(* IEC 61131-3 sources: Elmo_Master/Lasal_PRG/Elmo_EtherCAT_Test_4Axis/Class/ECAT_Slave_Base (part 2) *)

        sSDOData.Buffer.pSDOCallback$^VirtualBase^.NewInst(#UserPara, #UserResult);
      end_if;

//*******************************************************************************************************************************************************
  end_case;

END_FUNCTION

FUNCTION VIRTUAL GLOBAL ECAT_Slave_Base::ClassState::NewInst
	VAR_INPUT
		pPara 	: ^CmdStruct;
		pResult 	: ^Results;
	END_VAR
	VAR_OUTPUT
		ret_code 	: IprStates;
	END_VAR
  VAR
    TmpRetCode : iprStates;
    pNewElement   : t_pHWCGetHardwareDiagnosisOutDynExt;
    pTemp : ^void;
  END_VAR

  //Return with error if command is unknown or not supported
  ret_code := ERROR;

  case pPara^.uiCmd of

//**********************************************************************************************************************************************************
    ECAT_M_SET_SLAVE_INFO:

      pResult^.uiLng := 4;
      pResult^.aData[0]$DINT := ECAT_RETERR_CMD_VERSION;

      //Check version number
      if pPara^.aPara[0]$DINT = 1 then

        pResult^.uiLng := 8;
        pResult^.aData[0]$DINT := ECAT_RETERR_CMD_PARAMETER;
        pResult^.aData[4]$DINT := 1;  //Return version number

        pSlaveInfo := pPara^.aPara[1]$^t_st_eceni_slv_info;

        //Check for valid pointer
        if pSlaveInfo then

          ret_code := READY;

          //Show slave info data on server
          DeviceAdress  := pSlaveInfo^.physaddr;
          VendorID      := pSlaveInfo^.vendorid;
          SerialNo      := pSlaveInfo^.serialno;
          ProductCode   := pSlaveInfo^.productcode;
          RevisionNo    := pSlaveInfo^.revisionno;

          pResult^.aData[0]$DINT := ECATM_OK;

          if pSlaveInfo^.name then
            DeviceNameStr.WriteDataOff(udLen:=_StrLen(pSlaveInfo^.name), udOff:=0, pData:=pSlaveInfo^.name);
          else
            LogValue("@059A (ECAT_Slave_Base::ClassState::NewInst) Invalid name in Slave-info data of Slave 0x{0}",SlaveIndex);
          end_if;

          if pSlaveInfo^.productrev then
            ProductRevStr.WriteDataOff(udLen:=_StrLen(pSlaveInfo^.productrev), udOff:=0, pData:=pSlaveInfo^.productrev);
          else
            LogValue("@059B (ECAT_Slave_Base::ClassState::NewInst) Invalid product revision in Slave-info data of Slave 0x{0}",SlaveIndex);
          end_if;
        else

        end_if;
      else
        LogError("@059C (ECAT_Slave_Base::ClassState::NewInst) Unsupported NewInst version ECAT_M_SET_SLAVE_INFO");
        ret_code := ERROR;
      end_if;

//**********************************************************************************************************************************************************
    ECAT_M_GET_SLAVE_CYCIDX:

      pResult^.uiLng := 4;
      pResult^.aData[0]$DINT := ECAT_RETERR_CMD_VERSION;

      //Check version number
      if pPara^.aPara[0]$DINT = 1 then

        pResult^.uiLng := 8;
        pResult^.aData[4]$DINT := 1;  //Return version number

        pResult^.aData[0]$DINT := ECAT_RETERR_CMD_WRONG_SLV_STATE;
        if us_InitCnt >= 12 & ClassState = _ClassOk then

          pResult^.uiLng := 12;
          pResult^.aData[8]$DINT := to_dint(usCycIDX);
          pResult^.aData[0]$DINT := ECAT_RETOK;

          ret_code := READY;

//        else
//          // CYCIDX not set
        end_if;

      else
        LogError("@059D (ECAT_Slave_Base::ClassState::NewInst) Unsupported NewInst version ECAT_M_GET_SLAVE_CYCIDX");
        ret_code := ERROR;
      end_if;

//**********************************************************************************************************************************************************
    ECAT_M_EVENT_CALLBACK:
      pResult^.uiLng := 4;

      pResult^.aData[0]$DINT := ECAT_RETERR_CMD_VERSION;

      //Check version number
      if pPara^.aPara[0]$DINT = 1 then

        pResult^.uiLng := 8;
        pResult^.aData[0]$DINT := ECAT_RETOK;
        pResult^.aData[4]$DINT := 1;  //Return version number

        EvtCallBack(pPara^.aPara[1]$pVoid, pPara^.aPara[2]$^t_st_ecatm_evt, pPara^.aPara[3],pPara^.aPara[4]$UINT);

        ret_code := READY;
      else
        LogError("@059E (ECAT_Slave_Base::ClassState::NewInst) Unsupported NewInst version ECAT_M_EVENT_CALLBACK");
        ret_code := ERROR;
      end_if;

//**********************************************************************************************************************************************************
    ECAT_M_CHECK_SLAVE:

      pResult^.uiLng := 4;

      pResult^.aData[0]$DINT := ECAT_RETERR_CMD_VERSION;

      //Check version number
      if pPara^.aPara[0]$DINT = 1 then

        pResult^.uiLng := 8;
        pResult^.aData[4]$DINT := 1;  //Return version number

        pResult^.aData[0]$DINT := ECAT_RETERR;
        if CheckProductCode(udProductCodeToCheck:= pPara^.aPara[1]$UDINT
                          , udVendorIDToCheck   := pPara^.aPara[3]$UDINT) = TRUE then

          pResult^.aData[0]$DINT := ECAT_RETOK;
          ret_code := READY;

        end_if;

      else
        LogError("@059F (ECAT_Slave_Base::ClassState::NewInst) Unsupported NewInst version ECAT_M_CHECK_SLAVE");
        ret_code := ERROR;
      end_if;

//**********************************************************************************************************************************************************
    ECAT_M_CALL_INIT_MODULE:

      pResult^.uiLng := 4;

      pResult^.aData[0]$DINT := ECAT_RETERR_CMD_VERSION;

      //Check version number
      if pPara^.aPara[0]$DINT = 1 then

        pResult^.uiLng := 8;
        pResult^.aData[4]$DINT := 1;  //Return version number

        ret_code := InitModule(pPara^.aPara[1]$t_e_ECAT_STATE);

      else
        LogError("@05A1 (ECAT_Slave_Base::ClassState::NewInst) Unsupported NewInst version ECAT_M_CHECK_SLAVE");
        ret_code := ERROR;
      end_if;

//**********************************************************************************************************************************************************
    ECAT_M_SDO_CALLBACK:

      pResult^.uiLng := 4;

      pResult^.aData[0]$DINT := ECAT_RETERR_CMD_VERSION;

      //Check version number
      if pPara^.aPara[0]$DINT = 1 then

        pResult^.uiLng := 8;
        pResult^.aData[4]$DINT := 1;  //Return version number

        ret_code := READY;
        pResult^.aData[0]$DINT := ECAT_RETOK;

        ReceiveSDOResponse(sd_retval        := pPara^.aPara[1]
                         , bReadOrWriteSDO  := pPara^.aPara[2]$BOOL
                         , hIndex           := pPara^.aPara[3]$HINT
                         , hsSubIndex       := pPara^.aPara[4]$HSINT
                         , usLength         := pPara^.aPara[5]$USINT
                         , udErrorCode      := pPara^.aPara[6]$UDINT
                         );
      else
        LogError("@05A2 (ECAT_Slave_Base::ClassState::NewInst) Unsupported NewInst version ECAT_M_SDO_CALLBACK");
        ret_code := ERROR;
      end_if;

//**********************************************************************************************************************************************************
    ECAT_M_GET_HW_PATH:

      ret_code  := ERROR;
      pTemp     := NIL;

      //Check version
      pResult^.aData[0]$DINT  := ECAT_RETERR_CMD_VERSION;
      if (pPara^.aPara[0]$DINT = 2) then

        pTemp := GetPointer2ObjectPath(NIL);

        if pTemp then
          pResult^.aData[0]$DINT := ECAT_RETOK;
          ret_code := READY;
        else
          pResult^.aData[0]$DINT  := ECAT_RETERR;
        end_if;

        pResult^.uiLng := 14;
        pResult^.aData[4]$DINT    := 2; //Version
        pResult^.aData[8]$^void   := pTemp;
        pResult^.aData[12]$HSINT  := 0; // 0 This is Slave, Value is set by EtherCAT_Hub_Base
        pResult^.aData[13]$HINT   := 0; // 0 This is Slave, Value is set by EtherCAT_Hub_Base

      else
        // Version 1 is handled directly by Master Class
        // Passes on the NewInst command
        ret_code := toMaster.NewInst(pPara,pResult);
      end_if;

//**********************************************************************************************************************************************************
    ECAT_M_SET_CLASSSTATE:

      pResult^.uiLng := 4;

      pResult^.aData[0]$DINT := ECAT_RETERR_CMD_VERSION;

      //Check version number
      if pPara^.aPara[0]$DINT = 1 then

        pResult^.uiLng := 8;
        pResult^.aData[4]$DINT := 1;  //Return version number

        ret_code := READY;
        pResult^.aData[0]$DINT := ECAT_RETOK;

        ClassState := pPara^.aPara[1]$t_e_VaranErrors;
        Online     := pPara^.aPara[2]$DINT;
      else
        LogError("@084C (ECAT_Slave_Base::ClassState::NewInst) Unsupported NewInst version ECAT_M_SET_CLASSSTATE");
        ret_code := ERROR;
      end_if;

//**********************************************************************************************************************************************************
    ECAT_M_START_SDO:

      pResult^.uiLng := 4;

      pResult^.aData[0]$DINT := ECAT_RETERR_CMD_VERSION;

      //Check version number
      if pPara^.aPara[0]$DINT = 1 then

        pResult^.uiLng := 8;
        pResult^.aData[4]$DINT := 1;  //Return version number

        if pPara^.aPara[1] = 0 then
          ret_code := StartReadSDO( hIndex          := pPara^.aPara[2]$HINT
                                  , hsSubIndex      := pPara^.aPara[3]$HSINT
                                  , dCompleteAccess := pPara^.aPara[4]
                                  , pReadData       := pPara^.aPara[5]$^USINT
                                  , udMaxDataLength := pPara^.aPara[6]$UDINT
                                  , udTimeout       := pPara^.aPara[7]$UDINT
                                  , pCallback       := pPara^.aPara[8]$pVoid);
        else
          ret_code := StartWriteSDO(hIndex          := pPara^.aPara[2]$HINT
                                  , hsSubIndex      := pPara^.aPara[3]$HSINT
                                  , dCompleteAccess := pPara^.aPara[4]
                                  , pWriteData      := pPara^.aPara[5]$^USINT
                                  , udWriteLength   := pPara^.aPara[6]$UDINT
                                  , udTimeout       := pPara^.aPara[7]$UDINT
                                  , pCallback       := pPara^.aPara[8]$pVoid);
        end_if;

        if ret_code = READY then
          pResult^.aData[0]$DINT := ECAT_RETOK;
        elsif ret_code = BUSY then
          pResult^.aData[0]$DINT := ECAT_RETBUSY;
        else
          pResult^.aData[0]$DINT := ECAT_RETERR_CMD_PARAMETER;
        end_if;

      end_if;

//*********************************************************************************************************************************************************
    ECAT_M_START_ASYCOM:

      pResult^.uiLng := 4;

      pResult^.aData[0]$DINT := ECAT_RETERR_CMD_VERSION;

      //Check version number
      if pPara^.aPara[0]$DINT = 1 then

        pResult^.uiLng := 8;
        pResult^.aData[4]$DINT := 1;  //Return version number

        if pPara^.aPara[1] = 0 then // Read

          ret_code := StartAsyncComRead(Address     := pPara^.aPara[2]$HDINT
                                      , pReadData   := pPara^.aPara[3]$^USINT
                                      , DataLength  := pPara^.aPara[4]$UINT
                                      , udTimeout   := pPara^.aPara[5]$UDINT
                                      , pCallback   := pPara^.aPara[6]$pVoid);
        else  // Write

          ret_code := StartAsyncComWrite( Address       := pPara^.aPara[2]$HDINT
                                        , pWriteData    := pPara^.aPara[3]$^USINT
                                        , udWriteLength := pPara^.aPara[4]$UINT
                                        , udTimeout     := pPara^.aPara[5]$UDINT
                                        , pCallback     := pPara^.aPara[6]$pVoid);
        end_if;

        if ret_code = READY then
          pResult^.aData[0]$DINT := ECAT_RETOK;
        elsif ret_code = BUSY then
          pResult^.aData[0]$DINT := ECAT_RETBUSY;
        else
          pResult^.aData[0]$DINT := ECAT_RETERR_CMD_PARAMETER;
        end_if;

      end_if;

//*********************************************************************************************************************************************************
    ECAT_M_START_FOE:

      pResult^.uiLng := 4;

      pResult^.aData[0]$DINT := ECAT_RETERR_CMD_VERSION;

      //Check version number
      if pPara^.aPara[0]$DINT = 1 then

        pResult^.uiLng := 8;
        pResult^.aData[4]$DINT := 1;  //Return version number

        if pPara^.aPara[1] = 0 then // Read
          ret_code := StartFileRead(FileName      := pPara^.aPara[2]$^Char
                                  , PassWord      := pPara^.aPara[3]$UDINT
                                  , pFileBuffer   := pPara^.aPara[4]$pVoid
                                  , FileBufferSize:= pPara^.aPara[5]$UDINT
                                  , udTimeout     := pPara^.aPara[6]$UDINT
                                  , pCallback     := pPara^.aPara[7]$pVoid
                                  );
        elsif pPara^.aPara[1] = 1 then // Write
          ret_code := StartFileWrite( FileName  := pPara^.aPara[2]$^Char
                                    , PassWord  := pPara^.aPara[3]$UDINT
                                    , pFile     := pPara^.aPara[4]$pVoid
                                    , FileSize  := pPara^.aPara[5]$UDINT
                                    , udTimeout := pPara^.aPara[6]$UDINT
                                    , pCallback := pPara^.aPara[7]$pVoid
                                    );
        elsif pPara^.aPara[1] = -1 then // Abort
          ret_code := AbortFileAccess();
        else
          // Unkown
          ret_code := ERROR;
        end_if;

        if ret_code = READY then
          pResult^.aData[0]$DINT := ECAT_RETOK;
        elsif ret_code = BUSY then
          pResult^.aData[0]$DINT := ECAT_RETBUSY;
        else
          pResult^.aData[0]$DINT := ECAT_RETERR_CMD_PARAMETER;
        end_if;

      end_if;

//*********************************************************************************************************************************************************
    ECAT_M_START_SSC:

      pResult^.uiLng := 4;

      pResult^.aData[0]$DINT := ECAT_RETERR_CMD_VERSION;

      //Check version number
      if pPara^.aPara[0]$DINT = 1 then

        pResult^.uiLng := 8;
        pResult^.aData[4]$DINT := 1;  //Return version number

        if pPara^.aPara[1] = 0 then // Read

          ret_code := StartReadSoESSC(driveno         := pPara^.aPara[2]
                                    , elementflags    := pPara^.aPara[3]$USINT
                                    , idn             := pPara^.aPara[4]
                                    , pReadData       := pPara^.aPara[5]$^USINT
                                    , udMaxDataLength := pPara^.aPara[6]$UDINT
                                    , udTimeout       := pPara^.aPara[7]$UDINT
                                    , pCallback       := pPara^.aPara[8]$pVoid
                                    );
        else  // Write
          ret_code := StartWriteSoESSC( driveno       := pPara^.aPara[2]
                                      , elementflags  := pPara^.aPara[3]$USINT
                                      , idn           := pPara^.aPara[4]
                                      , pWriteData    := pPara^.aPara[5]$^USINT
                                      , udWriteLength := pPara^.aPara[6]$UDINT
                                      , udTimeout     := pPara^.aPara[7]$UDINT
                                      , pCallback     := pPara^.aPara[8]$pVoid
                                      );
        end_if;

        if ret_code = READY then
          pResult^.aData[0]$DINT := ECAT_RETOK;
        elsif ret_code = BUSY then
          pResult^.aData[0]$DINT := ECAT_RETBUSY;
        else
          pResult^.aData[0]$DINT := ECAT_RETERR_CMD_PARAMETER;
        end_if;

      end_if;

//*********************************************************************************************************************************************************
    CMD_GET_HARDWARE_TREE_ENTRY :

      //Set Errors
      ret_code := ERROR;
      pResult^.aData$t_HWCGetHardwareTreeEntryOut.retcode := _HWC_RETVAL_ERROR;
      pResult^.aData[0]$t_HWCGetHardwareTreeEntryOut.pStr_NextHardewareTreeEntry := NIL;

      if pObjectPath then
        //Copy Length of p_objectpath (is on 1st byte) on first byte of our array, length is 2 byte so set the 2nd byte manual
        a_HWTEntryStr[0] := pObjectPath^$USINT;
        a_HWTEntryStr[1] := 0;

        //a_HWTEntryStr + 2 because first 2 bytes are lenght, ObjectPath 1st byte is length, copy as long as the object path is
        _memcpy(ptr1:=#a_HWTEntryStr+2, ptr2:=pObjectPath+1, cntr:=a_HWTEntryStr[0]);

        //Return Hardware Tree Entry and set return codes
        pResult^.aData[0]$t_HWCGetHardwareTreeEntryOut.pStr_NextHardewareTreeEntry := #a_HWTEntryStr[0];
        ret_code := READY;
        pResult^.aData[0]$t_HWCGetHardwareTreeEntryOut.retcode := _HWC_RETVAL_OK_HWTSTR_RETURNED;

        // Compare Module string with passed string
        if pPara^.aPara[0]$t_HWCGetHardwareTreeEntryIn.pStr_LastHardewareTreeEntry then

          if pPara^.aPara[0]$t_HWCGetHardwareDiagnosisIn.pStr_HardewareTreeEntry$^USINT^ =
             pResult^.aData[0]$t_HWCGetHardwareTreeEntryOut.pStr_NextHardewareTreeEntry$^USINT^ then // Compare Length

            if _memcmp( ptr1:= pPara^.aPara[0]$t_HWCGetHardwareDiagnosisIn.pStr_HardewareTreeEntry // Compare Data
                      , ptr2:= pResult^.aData[0]$t_HWCGetHardwareTreeEntryOut.pStr_NextHardewareTreeEntry
                      , cntr:= pResult^.aData[0]$t_HWCGetHardwareTreeEntryOut.pStr_NextHardewareTreeEntry$^USINT^ + 2) = 0 then   // + 2 for 2 Byte Length

              pResult^.aData$t_HWCGetHardwareTreeEntryOut.retcode :=  _HWC_RETVAL_OK_MODULE_FOUND;
            end_if;
          end_if;
        end_if;
      end_if;

//**********************************************************************************************************************************************************
    CMD_GET_HARDWARE_DIAGNOSIS:

      pResult^.aData$t_HWCGetHardwareDiagnosisOut.retcode := _HWC_RETVAL_ERROR;
      ret_code := ERROR;

      //Return State and Device ID and set retcode ----------------------------------------------------------
      pResult^.aData$t_HWCGetHardwareDiagnosisOut.ClassState  := ClassState;
      pResult^.aData$t_HWCGetHardwareDiagnosisOut.ud_DeviceID := GetDeviceID();

      if ClassState = _NoHardware then
        pResult^.aData$t_HWCGetHardwareDiagnosisOut.retcode := _HWC_RETVAL_ERROR_NO_HARDWARE;
        return;
      elsif ClassState = _WrongHardware then
        pResult^.aData$t_HWCGetHardwareDiagnosisOut.retcode := _HWC_RETVAL_ERROR_WRONG_HARDWARE;
        return;
      elsif ClassState = _NoCalibDataFound then
        pResult^.aData$t_HWCGetHardwareDiagnosisOut.retcode := _HWC_RETVAL_ERROR_NO_CALIB_DATA_FOUND;
        return;
      elsif ClassState <> _ClassOk then
        pResult^.aData$t_HWCGetHardwareDiagnosisOut.retcode := _HWC_RETVAL_ERROR_NO_HARDWARE;
        return;
      end_if;

      //------------------------------------------------------------------------------------------------------

      if this <> p_this then
        //Reset statemachine
        eSDOSSW := _GetDeviceName;
        //Save This pointer
        p_this := this;

        // Reset Flags
        bDiagnosisDataAvailableFlags.HWVersion        := FALSE;
        bDiagnosisDataAvailableFlags.IdentityObject   := FALSE;
        bDiagnosisDataAvailableFlags.DeviceName       := FALSE;
        bDiagnosisDataAvailableFlags.SoftwareVersion  := FALSE;
      end_if;

      case eSDOSSW of

        //***********************************************************************************************************************************
        t_e_SDOSSW::_GetDeviceName:

          ret_code := BUSY;

          case eResponseStateHardwareTreeDiagnosis of
            //*****************************************************************************************
            t_e_ResponseStateSDO::_idle:

              TmpRetCode := StartReadSDO(hIndex          := ECAT_SB_INDEX_DEVICE_NAME
                                       , hsSubIndex      := ECAT_SB_SUBINDEX_DEVICE_NAME
                                       , dCompleteAccess := 0
                                       , pReadData       := #a_DeviceName[0]
                                       , udMaxDataLength := sizeof(a_DeviceName)
                                       , udTimeout       := ECAT_SB_DEFAULT_SDO_TIMEOUT
                                       , pCallback       := THIS
                                       );

              if TmpRetCode = READY then
                eResponseStateHardwareTreeDiagnosis := _wait;
                udSDOTimeout := ops.tAbsolute;

              elsif TmpRetCode = ERROR then
                ret_code := ERROR;
                eSDOSSW := _DataReady;
              end_if;

            //*****************************************************************************************
            t_e_ResponseStateSDO::_wait:

              //Timeout-Check
              if ((ops.tAbsolute - udSDOTimeout) > ECAT_SB_DEFAULT_SDO_TIMEOUT) then
                LogError("@02D1 (ECAT_Slave_Base::ClassState::NewInst) SDO Response timeout read state at HWT Diagnosis");
                ret_code := ERROR;
              end_if;

            //*****************************************************************************************
            t_e_ResponseStateSDO::_valid:

              eResponseStateHardwareTreeDiagnosis := t_e_ResponseStateSDO::_idle;

              //Check for an SDO error
              if sSDOData.sd_retval = 0 then
                eSDOSSW := _GetIdentityObject;
                bDiagnosisDataAvailableFlags.DeviceName := TRUE;
                pResult^.aData[0]$t_HWCGetHardwareDiagnosisOut.pStr_DeviceName  := (#a_DeviceName)$^CHAR;

              else
                ret_code := ERROR;
                //Error
                pResult^.aData[0]$t_HWCGetHardwareDiagnosisOut.retcode := _HWC_RETVAL_ERROR_ECAT_SDO_ACCESS_FAILED;
              end_if;

          end_case;

        //***********************************************************************************************************************************
        t_e_SDOSSW::_GetIdentityObject:

          ret_code := BUSY;

          case eResponseStateHardwareTreeDiagnosis of
            //*****************************************************************************************
            t_e_ResponseStateSDO::_idle:

              TmpRetCode := StartReadSDO(hIndex          := ECAT_SB_INDEX_IDENTITY_OBJECT
                                       , hsSubIndex      := ECAT_SB_SUBINDEX_IDENTITY_OBJECT
                                       , dCompleteAccess := 1
                                       , pReadData       := #s_IdentityObject[0]
                                       , udMaxDataLength := sizeof(s_IdentityObject)
                                       , udTimeout       := ECAT_SB_DEFAULT_SDO_TIMEOUT
                                       , pCallback       := THIS
                                       );

              if TmpRetCode = READY then
                eResponseStateHardwareTreeDiagnosis := _wait;
                udSDOTimeout := ops.tAbsolute;
              elsif TmpRetCode = ERROR then
                ret_code := ERROR;
                eSDOSSW := _DataReady;
              end_if;

            //*****************************************************************************************
            t_e_ResponseStateSDO::_wait:

              //Timeout-Check
              if ((ops.tAbsolute - udSDOTimeout) > ECAT_SB_DEFAULT_SDO_TIMEOUT) then
                LogError("@02D1 (ECAT_Slave_Base::ClassState::NewInst) SDO Response timeout read state at HWT Diagnosis");
                ret_code := ERROR;
              end_if;

            //*****************************************************************************************
            t_e_ResponseStateSDO::_valid:

              eResponseStateHardwareTreeDiagnosis := t_e_ResponseStateSDO::_idle;

              //Check for an SDO error
              if sSDOData.sd_retval = 0 then
                eSDOSSW := _GetSoftwareVersion;
                bDiagnosisDataAvailableFlags.IdentityObject := TRUE;
                pResult^.aData[0]$t_HWCGetHardwareDiagnosisOut.ud_VendorID := s_IdentityObject$t_s_IdentityObject.udVendorID;
                pResult^.aData[0]$t_HWCGetHardwareDiagnosisOut.ud_DeviceID := s_IdentityObject$t_s_IdentityObject.udProductCode;
              else
                ret_code := ERROR;
                //Error
                pResult^.aData[0]$t_HWCGetHardwareDiagnosisOut.retcode := _HWC_RETVAL_ERROR_ECAT_SDO_ACCESS_FAILED;
              end_if;

          end_case;
        //***********************************************************************************************************************************
        t_e_SDOSSW::_GetSoftwareVersion:

          ret_code := BUSY;

          case eResponseStateHardwareTreeDiagnosis of
            //*****************************************************************************************
            t_e_ResponseStateSDO::_idle:

              TmpRetCode := StartReadSDO(hIndex          := ECAT_SB_INDEX_SOFTWARE_VERSION
                                       , hsSubIndex      := ECAT_SB_SUBINDEX_SOFTWARE_VERSION
                                       , dCompleteAccess := 0
                                       , pReadData       := #a_FWVersion[0]
                                       , udMaxDataLength := sizeof(a_FWVersion)
                                       , udTimeout       := ECAT_SB_DEFAULT_SDO_TIMEOUT
                                       , pCallback       := THIS
                                       );

              if TmpRetCode = READY then
                eResponseStateHardwareTreeDiagnosis := _wait;
                udSDOTimeout := ops.tAbsolute;
              elsif TmpRetCode = ERROR then
                ret_code := ERROR;
                eSDOSSW := _DataReady;
              end_if;

            //*****************************************************************************************
            t_e_ResponseStateSDO::_wait:

              //Timeout-Check
              if ((ops.tAbsolute - udSDOTimeout) > ECAT_SB_DEFAULT_SDO_TIMEOUT) then
                LogError("@02D1 (ECAT_Slave_Base::ClassState::NewInst) SDO Response timeout read state at HWT Diagnosis");
                ret_code := ERROR;
              end_if;

            //*****************************************************************************************
            t_e_ResponseStateSDO::_valid:

              eResponseStateHardwareTreeDiagnosis := t_e_ResponseStateSDO::_idle;

              //Check for an SDO error
              if sSDOData.sd_retval = 0 then
                eSDOSSW := _GetHardwareVersion;
                bDiagnosisDataAvailableFlags.SoftwareVersion := TRUE;
                pResult^.aData[0]$t_HWCGetHardwareDiagnosisOut.pStr_FWVersion  := (#a_FWVersion)$^CHAR;

              else
                ret_code := ERROR;
                //Error
                pResult^.aData[0]$t_HWCGetHardwareDiagnosisOut.retcode := _HWC_RETVAL_ERROR_ECAT_SDO_ACCESS_FAILED;
              end_if;
          end_case;

        //***********************************************************************************************************************************
        t_e_SDOSSW::_GetHardwareVersion:

          ret_code := BUSY;

          case eResponseStateHardwareTreeDiagnosis of
            //*****************************************************************************************
            t_e_ResponseStateSDO::_idle:

              TmpRetCode := StartReadSDO(hIndex          := ECAT_SB_INDEX_HARDWARE_VERSION
                                       , hsSubIndex      := ECAT_SB_SUBINDEX_HARDWARE_VERSION
                                       , dCompleteAccess := 0
                                       , pReadData       := #a_HwVersion[0]
                                       , udMaxDataLength := sizeof(a_HwVersion)
                                       , udTimeout       := ECAT_SB_DEFAULT_SDO_TIMEOUT
                                       , pCallback       := THIS
                                       );

              if TmpRetCode = READY then
                eResponseStateHardwareTreeDiagnosis := _wait;
                udSDOTimeout := ops.tAbsolute;
              elsif TmpRetCode = ERROR then
                ret_code := ERROR;
                eSDOSSW := _DataReady;
              end_if;

            //*****************************************************************************************
            t_e_ResponseStateSDO::_wait:

              //Timeout-Check
              if ((ops.tAbsolute - udSDOTimeout) > ECAT_SB_DEFAULT_SDO_TIMEOUT) then
                LogError("@02D1 (ECAT_Slave_Base::ClassState::NewInst) SDO Response timeout read state at HWT Diagnosis");
                ret_code := ERROR;
              end_if;

            //*****************************************************************************************
            t_e_ResponseStateSDO::_valid:

              eResponseStateHardwareTreeDiagnosis := t_e_ResponseStateSDO::_idle;

              //Check for an SDO error
              if sSDOData.sd_retval = 0 then
                eSDOSSW := _DataReady;
                bDiagnosisDataAvailableFlags.HWVersion := TRUE;
              else
                ret_code := ERROR;
                //Error
                pResult^.aData[0]$t_HWCGetHardwareDiagnosisOut.retcode := _HWC_RETVAL_ERROR_ECAT_SDO_ACCESS_FAILED;
              end_if;
          end_case;

        //***********************************************************************************************************************************
        t_e_SDOSSW::_DataReady:

          //Not available for EtherCAT modules
          pResult^.aData[0]$t_HWCGetHardwareDiagnosisOut.pStr_VendorName := NIL;
          pResult^.aData[0]$t_HWCGetHardwareDiagnosisOut.pStr_OrderingNo := NIL;

          // first free the old then create the memory (linked list) for the additional information
          if pAdditionalDiagInfo then
            HwDiagFreeDynExtList(pList:=pAdditionalDiagInfo);
          end_if;
          pAdditionalDiagInfo      := NIL;

          //Data which is already available in HWK
          pResult^.aData[0]$t_HWCGetHardwareDiagnosisOut.ud_Place := SlaveIndex;

          if bDiagnosisDataAvailableFlags.DeviceName then
            pResult^.aData[0]$t_HWCGetHardwareDiagnosisOut.pStr_DeviceName  := (#a_DeviceName)$^CHAR;
          end_if;

          if bDiagnosisDataAvailableFlags.SoftwareVersion then
            pResult^.aData[0]$t_HWCGetHardwareDiagnosisOut.pStr_FWVersion  := (#a_FWVersion)$^CHAR;
          end_if;

          if bDiagnosisDataAvailableFlags.IdentityObject then
            pResult^.aData[0]$t_HWCGetHardwareDiagnosisOut.ud_VendorID := s_IdentityObject$t_s_IdentityObject.udVendorID;
            pResult^.aData[0]$t_HWCGetHardwareDiagnosisOut.ud_DeviceID := s_IdentityObject$t_s_IdentityObject.udProductCode;

            // add the serialnumber
            pNewElement := HwDiagAddDynExt2List(ppList:=#pAdditionalDiagInfo, EntryID:=_HWC_DIAG_ID_UDINT_SERIAL_NUMBER, udVersion:=1, udDataLength:=sizeof(t_s_IdentityObject.udSerialnumber));

            if pNewElement then
              (pNewElement$^HDINT + sizeof(t_HWCGetHardwareDiagnosisOutDynExt))^ := s_IdentityObject$t_s_IdentityObject.udSerialnumber;
            end_if;

          end_if;

          if bDiagnosisDataAvailableFlags.HWVersion then
          // add the hardware version
            pNewElement := HwDiagAddDynExt2List(ppList:=#pAdditionalDiagInfo, EntryID:=_HWC_DIAG_ID_STRING_HARDWARE_VERSION, udVersion:=1, udDataLength:=_strlen(src:=#a_HWVersion[0]));

            if pNewElement then
              // add the data in the reserved memory
              _strcpy(dest:=(pNewElement$^HDINT + sizeof(t_HWCGetHardwareDiagnosisOutDynExt))$^CHAR, src:=#a_HWVersion[0]);
            end_if;
          end_if;

          pResult^.aData[0]$t_HWCGetHardwareDiagnosisOut.p_DynExtList := pAdditionalDiagInfo;

          ret_code := READY;
          pResult^.aData[0]$t_HWCGetHardwareDiagnosisOut.retcode := _HWC_RETVAL_OK;

      end_case;

//**********************************************************************************************************************************************************
    ECAT_SB_GET_SLVIDX:
      pResult^.uiLng := 8;

      pResult^.aData[0]$DINT := 1;  //Return version number
      pResult^.aData[4]$DINT := ECAT_RETERR_CMD_VERSION;

      //Check version number
      if pPara^.aPara[0]$DINT = 1 then

        pResult^.uiLng := 12;
        pResult^.aData[4]$DINT := ECAT_RETOK;
        pResult^.aData[8]$UDINT := SlaveIndex;

        ret_code := READY;
      end_if;

//**********************************************************************************************************************************************************
    else
      // Passes on the NewInst command
      ret_code := toMaster.NewInst(pPara,pResult);
  end_case;

END_FUNCTION

FUNCTION __CDECL ECAT_Slave_Base::EvtCallBack
  VAR_INPUT
    pecatmhdl       : pVoid;
    evt             : ^t_st_ecatm_evt;
    EventType       : DINT;
    uiCallbackInfo  : UINT;
  END_VAR

  case evt^.evtcode of

//*******************************************************************************************************************************************************
  	ECATM_EVTC_SLV_STATE_CHANGE:

      EvtCallBackStateChange(evt^.arg3$UDINT);

//*******************************************************************************************************************************************************
  	ECATM_EVTC_SLV_TRANS_FAILED:

      EvtCallBackStateChange(evt^.arg3$UDINT);

      ClassState := _ClientNotready;
      Online     := 0;

      if uiCallbackInfo = LSL_ECATM_ACYCLIC_TASK then
        LogValue("@05A3 (ECAT_Slave_Base::EvtCallBack) ECATM_EVTC_SLV_TRANS_FAILED error code = 0x{0}", evt^.arg4$UDINT);
      else
        bd_LogRtMessagesInCy.PostIt.EvtCallSlvTransFailed := TRUE;
        bd_LogRtMessagesInCy.aLogValue1[0]                := evt^.arg4$UDINT;
      end_if;

//*******************************************************************************************************************************************************
  	ECATM_EVTC_SLV_ACKERR_FAILED:

//*******************************************************************************************************************************************************
  	ECATM_EVTC_INITC_RCV_TMO:

      ClassState := _ClientNotready;
      Online     := 0;
      //Logging is done in master

//*******************************************************************************************************************************************************
  	ECATM_EVTC_INITC_VALID_WKC:

      ClassState := _ClientNotready;
      Online     := 0;
      //Logging is done in master

//*******************************************************************************************************************************************************
  	ECATM_EVTC_INITC_VALID_LEN:

      ClassState := _ClientNotready;
      Online     := 0;
      //Logging is done in master

//*******************************************************************************************************************************************************
  	ECATM_EVTC_INITC_VALID_DATA:

      ClassState := _ClientNotready;
      Online     := 0;
      //Logging is done in master

//*******************************************************************************************************************************************************
  	ECATM_EVTC_SUP_SLV_STATE_CHG:

      EvtCallBackStateChange(evt^.arg3$UDINT);

//*******************************************************************************************************************************************************
  	ECATM_EVTC_SUP_SLV_ALSTATUS_CHG:

      // arg2 is correct, compare debug log in ECAT_Master_Base::EvtCallBack -> ECATM_EVTC_SUP_SLV_ALSTATUS_CHG
      EvtCallBackStateChange(evt^.arg2$UDINT);

//*******************************************************************************************************************************************************
    ECATM_EVTC_SUP_SLV_COMM_CHG:

      EvtCallBackStateChange(evt^.arg3$UDINT);

  end_case;

END_FUNCTION

FUNCTION VIRTUAL ECAT_Slave_Base::EvtCallBackStateChange
	VAR_INPUT
		NewEtherCATState 	: UDINT;
	END_VAR
  VAR
  	retcode : DINT;
  END_VAR

  //Get slave status information
  retcode := OS_ECATM_SLV_GET_STATUS(pECAT, ecatmhdl, SlaveIndex, #sSlaveState);

  if retcode = ECATM_OK then
    AL_StatusCode := sSlaveState.alstatuscode;
  end_if;

#ifdef ECAT_DEBUG_EVENT_CALLBACKS
  if retcode = 0 then
    LogValue(pString:="ECAT-DEBUG: (ECAT_Slave_Base::EvtCallBackStateChange) CurrState: 0x{0}, ExpectedState: 0x{1} ", Value:= sSlaveState.curstate, Value2 := sSlaveState.expstate);
    LogValue(pString:="ECAT-DEBUG: (ECAT_Slave_Base::EvtCallBackStateChange) alstatuscode: 0x{0}, flags: 0x{1} ", Value:= sSlaveState.alstatuscode, Value2 := sSlaveState.flags);
  end_if;
#endif

  EtherCATState$UDINT := (NewEtherCATState AND 16#0F);  //Only show

  SlaveState          := NewEtherCATState;

  if (EtherCATState = ECAT_STATE_OP) & (ClassState = _ClassOk) then
    Online := 1;
  else
    Online := 0;
  end_if;

END_FUNCTION

FUNCTION VIRTUAL GLOBAL ECAT_Slave_Base::GetInitModuleFlags
	VAR_OUTPUT
		bdInitModuleFlags 	: BDINT;
	END_VAR

  // define in derivation which flags are used

// like this (flags see ecat_master_base.h)
//  bdInitModuleFlags := ECAT_INIT_MODULE_CALL_INIT OR ECAT_INIT_MODULE_CALL_PREOP OR ECAT_INIT_MODULE_CALL_SAFEOP;

  bdInitModuleFlags := ECAT_INIT_MODULE_NO_CALL;

END_FUNCTION

#pragma warning(disable:73);
FUNCTION VIRTUAL ECAT_Slave_Base::ReceiveSDOResponse
	VAR_INPUT
		sd_retval 	: DINT;
		bReadOrWriteSDO 	: BOOL;
		hIndex 	: HINT;
		hsSubIndex 	: HSINT;
		usLength 	: USINT;
		udErrorCode 	: UDINT;
	END_VAR

  sSDOData.sd_retval := sd_retval;

  if eResponseStateHardwareTreeDiagnosis = _wait then
    eResponseStateHardwareTreeDiagnosis := _valid;
  end_if;

END_FUNCTION

FUNCTION VIRTUAL ECAT_Slave_Base::ReceiveAsyComResponse
	VAR_INPUT
		sd_retval 	: DINT;
		bReadOrWriteSDO 	: BOOL;
		hIndex 	: HINT;
		hsSubIndex 	: HSINT;
		usLength 	: USINT;
		udErrorCode 	: UDINT;
	END_VAR

  sAsyncComData.sd_retval := sd_retval;

END_FUNCTION

#pragma warning(default:73);

FUNCTION VIRTUAL GLOBAL ECAT_Slave_Base::ConnectEvent

  // overwrite this, if initmodule is used, so _NotInitialized can be shown during initialisation
  ClassState      := _ClassOk;

  // Reset SDO Handling
  sSDOData.bSDODataValid := FALSE;
  sigclib_atomic_setU32(pValue:=#sSDOData.udIsSDOActive, value:=ECAT_SB_SDO_FREE);
  // Clear Pipe
  if sSDOData.pPipe then

    while cPipe_Get(pd:=#sSDOData.Buffer, p:=sSDOData.pPipe) = 1 do
    end_while;

  end_if;

  sAsyncComData.bSDODataValid := FALSE;
  sigclib_atomic_setU32(pValue:=#sAsyncComData.udIsSDOActive, value:=ECAT_SB_SDO_FREE);
  // Clear Pipe
  if sAsyncComData.pPipe then

    while cPipe_Get(pd:=#sAsyncComData.Buffer, p:=sAsyncComData.pPipe) = 1 do
    end_while;

  end_if;

  // Reset FoE Handling
  sFoEData.bFoEDataValid := FALSE;
  sigclib_atomic_setU32(pValue:=#sFoEData.udIsFoEActive, value:=ECAT_SB_SDO_FREE);

  // Reset SSC Handling
  sSSCData.bSSCDataValid := FALSE;
  sigclib_atomic_setU32(pValue:=#sSSCData.udIsSSCActive, value:=ECAT_SB_SDO_FREE);
  // Clear Pipe
  if sSSCData.pPipe then

    while cPipe_Get(pd:=#sSSCData.Buffer, p:=sSSCData.pPipe) = 1 do
    end_while;

  end_if;

END_FUNCTION

FUNCTION VIRTUAL GLOBAL ECAT_Slave_Base::DisconnectEvent

  // at the disconnect we can use directly the server
  ClassState    := _NoHardware;
  EtherCATState := ECAT_STATE_INIT;
  Online        := 0;

END_FUNCTION

#pragma warning(disable:73);
FUNCTION VIRTUAL GLOBAL ECAT_Slave_Base::InitModule
	VAR_INPUT
		MasterState 	: t_e_ECAT_STATE;
	END_VAR
	VAR_OUTPUT
		eModuleInitState 	: iprStates;
	END_VAR
#pragma warning(default:73);

  // should be overwritten by derivation to initialize the module via SDO in a state machine if necessary (return BUSY while initializing)
  eModuleInitState := READY;

END_FUNCTION

FUNCTION VIRTUAL GLOBAL ECAT_Slave_Base::GetPointer2ObjectPath
	VAR_INPUT
		pThisPointerOverride 	: pVirtualBase;
	END_VAR
	VAR_OUTPUT
		p_us_ObjectPath 	: ^USINT;
	END_VAR
  VAR
  	MyPara   : CmdStruct;
    MyResult : results;
    p_us_PreviousPath : ^USINT;
    PrevLength : UINT;
    i : DINT;
    pLastEscSeq : ^HSINT;
    LastEscSeq : HSINT;
    NextEscSeq : HSINT;
    NextPortNo : USINT;
  END_VAR

  if ( pObjectPath = NIL ) then

    MyPara.aPara[0]$DINT := 2; //Version of command

    MyPara.uiCmd := ECAT_M_GET_HW_PATH;
    if toMaster.NewInst(#MyPara, #MyResult) <> READY then
      if bd_SingleLog.GetHwPathFailed = FALSE then
        bd_SingleLog.GetHwPathFailed := TRUE;
        LogError("@05A4 (ECAT_Slave_Base::GetPointer2ObjectPath) [SL] Failed to get hardware path of preceding module");
      end_if;
    else

      // Find last escape Sequence
      p_us_PreviousPath := MyResult.aData[8]$^USINT;
      NextEscSeq  := MyResult.aData[12]$HSINT;
      NextPortNo  := MyResult.aData[13]$USINT;
      PrevLength  := p_us_PreviousPath^$UINT;

      LastEscSeq := 0;  // Last EscSeq in the HW Tree of the Previous Module
      pLastEscSeq := p_us_PreviousPath + p_us_PreviousPath^ + 1;
      for i := PrevLength to 0 by -1 do

        if (pLastEscSeq^ AND HWT_ESCAPE_SEQU) then
          LastEscSeq := pLastEscSeq^;
          exit;
        end_if;

        pLastEscSeq -= sizeof(HSINT);

      end_for;

      if (LastEscSeq = 0) | (LastEscSeq <> NextEscSeq) then
        // Insert NextEscSeq
        //alloc memory
        pObjectPath := ( ToStdLib.Malloc( size := p_us_PreviousPath^ + 1 + 2) )$^USINT; // + 1 Length HWPath, + 2 (EscSeq + PortNo)

        // Length of HW-Path is 1 Byte and does not include length itself
        ToStdLib.MemCpy ( dest   := pObjectPath
                        , source := p_us_PreviousPath
                        , size   := p_us_PreviousPath^ + 1  // Include length in memcpy
                        );

        // increase length
        pObjectPath^ += 2; // 1 Byte Escape sequence + 1 Byte Port
        (pObjectPath + pObjectPath^ - 1)^ := NextEscSeq;
        (pObjectPath + pObjectPath^ + 0)^ := NextPortNo;
      else
        // No change of EscSeq
        // alloc memory
        pObjectPath := ( ToStdLib.Malloc( size := p_us_PreviousPath^ + 1 + 1 ) )$^USINT;  // + 1 Length HWPath, + 1 PortNo

        // Length of HW-Path is 1 Byte and does not include length itself
        ToStdLib.MemCpy ( dest   := pObjectPath
                        , source := p_us_PreviousPath
                        , size   := p_us_PreviousPath^ + 1  // Include length in memcpy
                        );

        // increase length
        pObjectPath^ += 1; //1 Byte Port
        (pObjectPath + pObjectPath^)^ := NextPortNo;
      end_if;

      if pThisPointerOverride then
        //register object path in OS
        SetObjectThisp(pObjectPath:=pObjectPath, pthis:=pThisPointerOverride$UDINT);
      else
        //register object path in OS
        SetObjectThisp(pObjectPath:=pObjectPath, pthis:=this$UDINT);
      end_if;
    end_if;
  end_if;

  p_us_ObjectPath := pObjectPath;

END_FUNCTION

FUNCTION ECAT_Slave_Base::SetObjectThisp
	VAR_INPUT
		pObjectPath 	: ^USINT;
		pThis 	: UDINT;
	END_VAR
	VAR_OUTPUT
		dRetcode 	: DINT;
	END_VAR

  if ( pHardwareTree <> NIL ) then
    dRetcode := HWT_iSetObjectThisp(0,pObjectPath,pThis);
  else
    dRetcode := 0;
  end_if;

END_FUNCTION

FUNCTION ECAT_Slave_Base::GetObjectThisp
	VAR_INPUT
		pObjectPath 	: ^USINT;
	END_VAR
	VAR_OUTPUT
		pThis 	: UDINT;
	END_VAR

  if ( pHardwareTree <> NIL ) then
    pThis := HWT_iGetObjectThisp(0,pObjectPath);
  else
    pThis := 0;
  end_if;

END_FUNCTION

FUNCTION ECAT_Slave_Base::HwDiagFreeDynExtList
  VAR_INPUT
    pList 	: ^t_HWCGetHardwareDiagnosisOutDynExt;
  END_VAR
  VAR
    pHelp 	: ^t_HWCGetHardwareDiagnosisOutDynExt;
  END_VAR

  while pList do
    // remember the current entry
    pHelp := pList;

    // set plist to the next entry and free pHelp
    pList := pList^.p_Next;

    // free the current entry
    ToStdLib.Free(mptr:=pHelp);
  end_while;

END_FUNCTION

FUNCTION ECAT_Slave_Base::HwDiagAddDynExt2List
	VAR_INPUT
		ppList 	: ^t_pHWCGetHardwareDiagnosisOutDynExt;
		EntryID 	: t_HWCGetHardwareDiagnosisOutType;
		udVersion 	: UDINT;
		udDataLength 	: UDINT;
	END_VAR
	VAR_OUTPUT
		pNewElement 	: t_pHWCGetHardwareDiagnosisOutDynExt;
	END_VAR

  if ppList^ = NIL then
    ppList^$pVoid := ToStdLib.Malloc(size:=sizeof(t_HWCGetHardwareDiagnosisOutDynExt) + udDataLength);
    pNewElement := ppList^;
  else
    pNewElement := ppList^;
    while pNewElement^.p_Next <> NIL do
      pNewElement := pNewElement^.p_Next;
    end_while;
    pNewElement^.p_Next$pVoid := ToStdLib.Malloc(size:=sizeof(t_HWCGetHardwareDiagnosisOutDynExt) + udDataLength);
    pNewElement := pNewElement^.p_Next;
  end_if;

  if pNewElement <> NIL then
    // initialize the new memory
    pNewElement^.DiagID         := EntryID;
    pNewElement^.ud_Version     := udVersion;
    pNewElement^.p_Next         := NIL;
    pNewElement^.ud_DataLength  := udDataLength;

    if udDataLength then
      _memset(dest:=pNewElement + sizeof(t_HWCGetHardwareDiagnosisOutDynExt), usByte:=0, cntr:=udDataLength);
    end_if;
  end_if;

END_FUNCTION

FUNCTION VIRTUAL GLOBAL ECAT_Slave_Base::GetDeviceID
	VAR_OUTPUT
		output 	: UDINT;
	END_VAR

  //Overwrite in derived Classes
  output := HWC_INVALID_DEVICE_ID;

END_FUNCTION

FUNCTION ECAT_Slave_Base::CyclicAsyncComHandling
VAR
	UserPara  : CmdStruct;
  UserResult: Results;
  sd_retval : DINT;
  retcode : iprStates;
END_VAR

  case sAsyncComData.eSSW of

//*******************************************************************************************************************************************************
    0:  //Start SDO Request

        if (sAsyncComData.pPipe) &
           (sAsyncComData.bSDODataValid = FALSE) then

          if cPipe_Get(pd:=#sAsyncComData.Buffer, p:=sAsyncComData.pPipe) = 1 then

            sAsyncComData.bSDODataValid := TRUE;

          end_if;

        end_if;

        if sAsyncComData.bSDODataValid then

          if sAsyncComData.Buffer.bReadOrWriteCommand = FALSE then  // Read
            //Start SDO Upload via OS
            sd_retval := OS_ECATM_ASYNC_START( pECAT
                                             , ecatmhdl                           // ecatm : pVoid; (* Struct: _ecatm_hdl *)
                                             , ECATM_CMD_FPRD                     // configured physical read //cmd : USINT;
                                             , sAsyncComData.Buffer.Address       // addr : UDINT;
                                             , sAsyncComData.Buffer.pData$^USINT  // datasndrcv : ^USINT;
                                             , sAsyncComData.Buffer.uiLength      // size : UINT;
                                             , sAsyncComData.Buffer.udTimeout     // tmo_ms : UDINT;
                                             , #sAsyncComData.pSDOHandle          // asynchdlp : pVoid; (* Struct: _ecatm_asynchdl *)
                                             );
          else  // Write

            //Start SDO Upload via OS
            sd_retval := OS_ECATM_ASYNC_START( pECAT
                                             , ecatmhdl                           // ecatm : pVoid; (* Struct: _ecatm_hdl *)
                                             , ECATM_CMD_FPWR                     // configured physical write //cmd : USINT;
                                             , sAsyncComData.Buffer.Address       // addr : UDINT;
                                             , sAsyncComData.Buffer.pData$^USINT  // datasndrcv : ^USINT;
                                             , sAsyncComData.Buffer.uiLength      // size : UINT;
                                             , sAsyncComData.Buffer.udTimeout     // tmo_ms : UDINT;
                                             , #sAsyncComData.pSDOHandle          // asynchdlp : pVoid; (* Struct: _ecatm_asynchdl *)
                                             );

          end_if;

          if sd_retval = ECATM_OK then
            retcode := READY;

            sAsyncComData.eSSW := 1; //Go on, wait for answer in next step

          elsif sd_retval <> ECATM_EVTC_BUSY$DINT then
            retcode := ERROR;

            LogValue("@06B3 (ECAT_Slave_Base::CyclicAsyncComHandling) Async Com Error 0x{0} at Slave 0x{1} while starting Async Com",sd_retval$UDINT,SlaveIndex);

            // Reset before udIsSDOActive
            sAsyncComData.bSDODataValid    := FALSE;
            sigclib_atomic_setU32(pValue:=#sAsyncComData.udIsSDOActive, value:=ECAT_SB_SDO_FREE);

            if sAsyncComData.Buffer.pSDOCallback then
              UserPara.uiCmd           := ECAT_M_ASYCOM_CALLBACK;
              UserPara.aPara[0]$DINT   := 1;                                        //Version
              UserPara.aPara[1]$DINT   := sd_retval;                                //Return code
              UserPara.aPara[2]$BOOL   := sAsyncComData.Buffer.bReadOrWriteCommand; //Read or Write (0 ... Read , 1 ... Write)
              UserPara.aPara[3]        := to_dint(sAsyncComData.Buffer.Address);    //register adress
              UserPara.aPara[4]        := 0;                                        //0 (not used)
              UserPara.aPara[5]        := to_dint(sAsyncComData.Buffer.uiLength);   //Datalength
              UserPara.aPara[6]$UDINT  := sAsyncComData.uiWorkingCounter;           //Working counter (gets incremented with every successful read or write)

              sAsyncComData.Buffer.pSDOCallback$^VirtualBase^.NewInst(#UserPara, #UserResult);
            end_if;
          end_if;
        end_if;

//*******************************************************************************************************************************************************
    1:  //Receive SDO Response

      sd_retval := OS_ECATM_ASYNC_POLL(pECAT
                                     , ecatmhdl                         // ecatm : pVoid; (* Struct: _ecatm_hdl *)
                                     , sAsyncComData.pSDOHandle         // asynchdl : pVoid; (* Struct: _ecatm_asynchdl *)
                                     , #sAsyncComData.uiWorkingCounter  // wkc : ^UINT;
                                     );

      if sd_retval = ECATM_OK then
        retcode := READY;
      elsif sd_retval = ECATM_EVTC_BUSY$DINT then
        retcode := BUSY;
        return;
      else
        LogValue("@06B4 (ECAT_Slave_Base::CyclicAsyncComHandling) Async Com Error 0x{0} at Slave 0x{1} while receiving response for Address: 0x{2}",sd_retval$UDINT,SlaveIndex, to_udint(sAsyncComData.Buffer.Address) );
        retcode := ERROR;
      end_if;

      // Reset before udIsSDOActive
      sAsyncComData.bSDODataValid   := FALSE;
      sAsyncComData.pSDOHandle      := NIL;
      sigclib_atomic_setU32(pValue:=#sAsyncComData.udIsSDOActive, value:=ECAT_SB_SDO_FREE);

      sAsyncComData.eSSW := 0; //Reset SSW

      if sAsyncComData.Buffer.pSDOCallback then
        UserPara.uiCmd          := ECAT_M_ASYCOM_CALLBACK;
        UserPara.aPara[0]$DINT  := 1;                                         // Version
        UserPara.aPara[1]$DINT  := sd_retval;                                 // Return code
        UserPara.aPara[2]$BOOL  := sAsyncComData.Buffer.bReadOrWriteCommand;  // Read or Write (0 ... Read , 1 ... Write)
        UserPara.aPara[3]       := to_dint(sAsyncComData.Buffer.Address);     // register adress
        UserPara.aPara[4]       := 0;                                         // 0 (not used)
        UserPara.aPara[5]       := to_dint(sAsyncComData.Buffer.uiLength);    // Datalength
        UserPara.aPara[6]$UDINT := sAsyncComData.uiWorkingCounter;            // Working counter (gets incremented with every successful read or write)

        sAsyncComData.Buffer.pSDOCallback$^VirtualBase^.NewInst(#UserPara, #UserResult);
      end_if;

//*******************************************************************************************************************************************************
  end_case;

END_FUNCTION

FUNCTION VIRTUAL ECAT_Slave_Base::InitSDOBuffers

  // Init SDO Buffers
  NoSDOBuffer := NoSDOBuffer.Read();

  sSDOData.pPipe := NIL;
  if NoSDOBuffer >= 1 then

    sSDOData.pPipe := cPipe_CTor(record_size:=sizeof(t_s_SDOBufferEntry), record_no:=NoSDOBuffer$UDINT);

    if sSDOData.pPipe = NIL then
      ClassState := _MemoryFault;
      LogError("@0926 (ECAT_Slave_Base::InitSDOBuffers) Failed to allocate memory for SDO-Buffer-pipe");
      EtherCATState := ECAT_STATE_NONE;
      return;
    end_if;

  end_if;

  NoAsyncBuffer := NoAsyncBuffer.Read();

  if NoAsyncBuffer >= 1 then

    sAsyncComData.pPipe := cPipe_CTor(record_size:=sizeof(t_s_AsyncBufferEntry), record_no:=NoAsyncBuffer$UDINT);

    if sAsyncComData.pPipe = NIL then
      ClassState := _MemoryFault;
      LogError("@0927 (ECAT_Slave_Base::InitSDOBuffers) Failed to allocate memory for AsyncComData-Buffer-pipe");
      EtherCATState := ECAT_STATE_NONE;
      return;
    end_if;

  end_if;

  NoSSCBuffer := NoSSCBuffer.Read();

  if NoSSCBuffer >= 1 then

    if (pECAT^.version < ECATM_CIL_SOE_SUPPORT) then
      NoSSCBuffer := 0;
      ClassState := _InvalidConfguration;
      LogError("@0928 (ECAT_Slave_Base::InitSDOBuffers) SSC is not suppored by current OS!");
      EtherCATState := ECAT_STATE_NONE;
      return;
    else

      sSSCData.pPipe := cPipe_CTor(record_size:=sizeof(t_s_SoESSCBufferEntry), record_no:=NoSSCBuffer$UDINT);

      if sSSCData.pPipe = NIL then
        ClassState := _MemoryFault;
        LogError("@0929 (ECAT_Slave_Base::InitSDOBuffers) Failed to allocate memory for SSC-Buffer-pipe");
        EtherCATState := ECAT_STATE_NONE;
        return;
      end_if;

    end_if;

  end_if;

END_FUNCTION

FUNCTION VIRTUAL GLOBAL ECAT_Slave_Base::StartFileWrite
	VAR_INPUT
		FileName 	: ^Char;
		PassWord 	: UDINT;
		pFile 	: pVoid;
		FileSize 	: UDINT;
		udTimeout 	: UDINT;
		pCallback 	: pVoid;
	END_VAR
	VAR_OUTPUT
		retcode 	: iprStates;
	END_VAR

  //Mailbox communication is available when State is Pre-Op or higher
  if EtherCATState < ECAT_STATE_PREOP then
    retcode := ERROR;
    return;
  end_if;

  //Check input parameters
  if (FileName = NIL) |
     (pFile = NIL)    |
     (FileSize = 0) then
    retcode := ERROR;
    return;
  end_if;

  if pCallback = NIL then
    retcode := ERROR;
    return;
  end_if;

  retcode := BUSY;
  // Check if currently a FoE is active, if not get lock on variables
  if (sigclib_atomic_cmpxchgU32(pValue:= #sFoEData.udIsFoEActive, cmpVal:=ECAT_SB_SDO_FREE, newVal:=ECAT_SB_SDO_LOCK) = ECAT_SB_SDO_FREE) then

    // Copy data to variables
    sFoEData.Buffer.ReadWriteAbortFoE := 1; //write
    sFoEData.Buffer.FileName          := FileName;
    sFoEData.Buffer.PassWord          := PassWord;
    sFoEData.Buffer.pFile             := pFile;
    sFoEData.Buffer.FileSize          := FileSize;
    sFoEData.Buffer.udTimeout         := udTimeout;
    sFoEData.Buffer.pFoECallback      := pCallback;

    sFoEData.eSSW             := t_e_FoESSW::_Idle;

    // Set when all other data is set
    sFoEData.bFoEDataValid    := TRUE;

    retcode := READY;

  end_if;
END_FUNCTION

FUNCTION VIRTUAL GLOBAL ECAT_Slave_Base::StartFileRead
	VAR_INPUT
		FileName        : ^Char;
		PassWord        : UDINT;
		pFileBuffer     : pVoid;
    FileBufferSize  : UDINT;
		udTimeout       : UDINT;
		pCallback       : pVoid;
	END_VAR
	VAR_OUTPUT
		retcode 	: iprStates;
	END_VAR

  //Mailbox communication is available when State is Pre-Op or higher
  if EtherCATState < ECAT_STATE_PREOP then
    retcode := ERROR;
    return;
  end_if;

  //Check input parameters
  if (FileName = NIL)     |
     (pFileBuffer = NIL)  |
     (FileBufferSize = 0) then
    retcode := ERROR;
    return;
  end_if;

  if pCallback = NIL then
    retcode := ERROR;
    return;
  end_if;

  //Check if currently a FoE is active
  retcode := BUSY;

  // Check if currently a FoE is active, if not get lock on variables
  if (sigclib_atomic_cmpxchgU32(pValue:= #sFoEData.udIsFoEActive, cmpVal:=ECAT_SB_SDO_FREE, newVal:=ECAT_SB_SDO_LOCK) = ECAT_SB_SDO_FREE) then

    // Copy data to variables
    sFoEData.Buffer.ReadWriteAbortFoE := 0; //Read
    sFoEData.Buffer.FileName          := FileName;
    sFoEData.Buffer.PassWord          := PassWord;
    sFoEData.Buffer.pFile             := pFileBuffer;
    sFoEData.Buffer.FileSize          := FileBufferSize;
    sFoEData.Buffer.udTimeout         := udTimeout;
    sFoEData.Buffer.pFoECallback      := pCallback;

    sFoEData.eSSW             := t_e_FoESSW::_Idle;

    // Set when all other data is set
    sFoEData.bFoEDataValid    := TRUE;

    retcode := READY;

  end_if;

END_FUNCTION

FUNCTION VIRTUAL GLOBAL ECAT_Slave_Base::AbortFileAccess
	VAR_OUTPUT
		retcode 	: iprStates;
	END_VAR

  retcode := BUSY;

  if (sigclib_atomic_cmpxchgU32(pValue:= #sFoEData.udIsFoEActive, cmpVal:=ECAT_SB_SDO_FREE, newVal:=ECAT_SB_SDO_LOCK) = ECAT_SB_SDO_FREE) then

    // No File acces was active, nothing to to.
    retcode := READY;
    sigclib_atomic_setU32(pValue:=#sFoEData.udIsFoEActive, value:=ECAT_SB_SDO_FREE);

  else

    sFoEData.bAbortAccess := TRUE;

  end_if;

END_FUNCTION

FUNCTION ECAT_Slave_Base::CyclicFoEHandling

  if sFoEData.bAbortAccess then

    sFoEData.bAbortAccess := FALSE;

    case sFoEData.eSSW of

      t_e_FoESSW::_Idle,          //Start FoE Request
      t_e_FoESSW::_StartReadFile,
      t_e_FoESSW::_StartWriteFile:
        // File access has not been started yet
        // Set Values that are passed by callback
        sFoEData.sd_retval := ECATM_OK;
        sFoEData.Buffer.FileName    := NIL;  // Clear string, may be old
        sFoEData.FileSizeTransferred := 0;
        _memset(dest:=#sFoEData.FoEStatus, usByte:=0, cntr:=sizeof(sFoEData.FoEStatus));  // Reset Status as it is used in callback and my not be filled in error

        sFoEData.Buffer.ReadWriteAbortFoE := -1;  // Set to -1 for abort callback
        sFoEData.eSSW := t_e_FoESSW::_Finish; // FoE Was not active, Nothing to do, set Finish for callback info

      t_e_FoESSW::_ReadFile,
      t_e_FoESSW::_WriteFile:

        // File access has is active => abort
        sFoEData.Buffer.ReadWriteAbortFoE := -1;  // Set to -1 for abort callback
        sFoEData.eSSW := t_e_FoESSW::_AbortFileAccess; // FoE is active, set SSW to abort

      t_e_FoESSW::_Finish,
      t_e_FoESSW::_Error:

        // File access already done, nothing todo

    end_case;
  end_if;

  case sFoEData.eSSW of

//*******************************************************************************************************************************************************
   t_e_FoESSW::_Idle:  //Start FoE Request

        if sFoEData.bFoEDataValid then

          if sFoEData.Buffer.ReadWriteAbortFoE = 0 then  // Read
            sFoEData.eSSW := t_e_FoESSW::_StartReadFile;
          elsif sFoEData.Buffer.ReadWriteAbortFoE > 0 then  // Write
            sFoEData.eSSW := t_e_FoESSW::_StartWriteFile;
          else // Abort < 0

          end_if;

        end_if;

//*******************************************************************************************************************************************************
    t_e_FoESSW::_StartReadFile:

        //Start FoE Upload via OS
        sFoEData.sd_retval := OS_ECATM_FOE_UPL_START( pECAT
                                                    , ecatmhdl                  // ecatm     : pVoid; (* Struct: _ecatm_hdl *)
                                                    , SlaveIndex                // slvidx    : UDINT;
                                                    , sFoEData.Buffer.FileName  // file      : ^char; (* const *)
                                                    , sFoEData.Buffer.PassWord  // password  : UDINT;
                                                    , sFoEData.Buffer.udTimeout // tmo_ms    : UDINT;
                                                    , #sFoEData.BlockSize       // blocksize : ^UDINT;
                                                    , #sFoEData.pFoEHandle      // trfhdlp   : pVoid; (* Struct: pointer to _ecatm_foe_trfhdl *)
                                                    );

        if sFoEData.sd_retval = ECATM_OK then

          sFoEData.eSSW := _ReadFile; //Go on, wait for answer in next step
          sFoEData.FileSizeTransferred := 0;
          _memset(dest:=#sFoEData.FoEStatus, usByte:=0, cntr:=sizeof(sFoEData.FoEStatus));  // Reset Status as it is used in callback and my not be filled in error

          if sFoEData.BlockSize > sFoEData.RdBlockBufferSize then

            if sFoEData.pRdBlockBuffer then

              sFoEData.pRdBlockBuffer     := toStdLib.ReAlloc(mptr:=sFoEData.pRdBlockBuffer, newsize:=sFoEData.BlockSize);
              sFoEData.RdBlockBufferSize  := sFoEData.BlockSize;

            else

              sFoEData.pRdBlockBuffer     := toStdLib.Malloc(size:=sFoEData.BlockSize);
              sFoEData.RdBlockBufferSize  := sFoEData.BlockSize;

            end_if;

            if sFoEData.pRdBlockBuffer = NIL then

              sFoEData.RdBlockBufferSize := 0;
              HWC_LogPrintf(pThis:=this, format:="@092A (ECAT_Slave_Base::CyclicFoEHandling) Failed to allocate memory for File read buffer.");
              sFoEData.eSSW := t_e_FoESSW::_Error;

            end_if;

          end_if;

        elsif sFoEData.sd_retval <> ECATM_EVTC_BUSY$DINT then

          sFoEData.eSSW := t_e_FoESSW::_Error;
          HWC_LogPrintf(pThis:=this, format:="@092B (ECAT_Slave_Base::CyclicFoEHandling) Call OS_ECATM_FOE_UPL_START returned %d.", p0:=#sFoEData.sd_retval);

        end_if;

//*******************************************************************************************************************************************************
    t_e_FoESSW::_ReadFile:

        sFoEData.sd_retval := OS_ECATM_FOE_UPL_POLL(pECAT
                                                  , ecatmhdl                        // ecatm   : pVoid; (* Struct: _ecatm_hdl *)
                                                  , sFoEData.pFoEHandle             // trfhdlp : pVoid; (* Struct: _ecatm_foe_trfhdl *)
                                                  , sFoEData.pRdBlockBuffer$^USINT  // data    : ^USINT;
                                                  , #sFoEData.FoEStatus             // status  : pVoid; (* Struct: pointer to _ecatm_foe_status *)
                                                  );

        if sFoEData.sd_retval = ECATM_OK then

          case sFoEData.FoEStatus.state of

            ECATM_FOE_IDLE:           // transfer completed; handle freed

              sFoEData.eSSW := t_e_FoESSW::_Finish; //Go on

            ECATM_FOE_DATA_READY:     // data chunk filled

              // Check if chunck fits in dest. pointer
              if ((sFoEData.FileSizeTransferred + sFoEData.FoEStatus.lastsize$UDINT) <= sFoEData.Buffer.FileSize) then

                // Copy chunk
                _memcpy(ptr1:=sFoEData.Buffer.pFile + sFoEData.FileSizeTransferred, ptr2:=sFoEData.pRdBlockBuffer, cntr:=sFoEData.FoEStatus.lastsize$UDINT);
                sFoEData.FileSizeTransferred += sFoEData.FoEStatus.lastsize$UDINT;

                // Send Update to user with new sFoEData.FileSizeTransferred
                SendFOECallback(FOEState:=BUSY);

              else

                sFoEData.eSSW := t_e_FoESSW::_AbortFileAccessError;  // Abort FoE Current File Access
                sFoEData.sd_retval := ECATM_EVTC_ERR_BUFSIZE;

                sFoEData.Buffer.ReadWriteAbortFoE := -1;  // Set to -1 for abort callback
                sFoEData.FileSizeTransferred += sFoEData.FoEStatus.lastsize$UDINT; // Only for callback
                HWC_LogPrintf(pThis:=this, format:="@092D (ECAT_Slave_Base::CyclicFoEHandling) Receive buffer for file %d is to small. At least %v Bytes are required.", p0:=#sFoEData.Buffer.FileSize, p1:=#sFoEData.FileSizeTransferred);
              end_if;

            ECATM_FOE_WAIT_BUFFER:    // buffer transferred

              // Nothing to do

            ECATM_FOE_BUSY:           // FoE transfer is busy

              // Nothing to do

            ECATM_FOE_ERROR:          // FoE transfer failed; handle freed

              sFoEData.eSSW := t_e_FoESSW::_Error;
              if sFoEData.FoEStatus.error_str[0] then
                sFoEData.FoEStatus.error_str[ECATM_FOE_MAXSTRLEN-1] := 0;   //Ensure 0 Terminaton
                HWC_LogPrintf(pThis:=this, format:="@092E (ECAT_Slave_Base::CyclicFoEHandling) Call OS_ECATM_FOE_UPL_POLL returned ErrorCode; %V2, Error Msg: %s", p0:=#sFoEData.FoEStatus.error_code, p1:=#sFoEData.FoEStatus.error_str[0]);
              else
                HWC_LogPrintf(pThis:=this, format:="@092E (ECAT_Slave_Base::CyclicFoEHandling) Call OS_ECATM_FOE_UPL_POLL returned ErrorCode %V2", p0:=#sFoEData.FoEStatus.error_code);
              end_if;

          end_case;

        else
          sFoEData.eSSW := t_e_FoESSW::_Error;
          HWC_LogPrintf(pThis:=this, format:="@092E (ECAT_Slave_Base::CyclicFoEHandling) Call OS_ECATM_FOE_UPL_POLL returned %d", p0:=#sFoEData.sd_retval);
        end_if;

//*******************************************************************************************************************************************************
    t_e_FoESSW::_StartWriteFile:

        sFoEData.sd_retval := OS_ECATM_FOE_DLD_START( pECAT
                                                    , ecatmhdl                  // ecatm     : pVoid; (* Struct: _ecatm_hdl *)
                                                    , SlaveIndex                // slvidx    : UDINT;
                                                    , sFoEData.Buffer.FileName  // file      : ^char; (* const *)
                                                    , sFoEData.Buffer.PassWord  // password  : UDINT;
                                                    , sFoEData.Buffer.udTimeout // tmo_ms    : UDINT;
                                                    , #sFoEData.BlockSize       // blocksize : ^UDINT;
                                                    , #sFoEData.pFoEHandle      // trfhdlp   : pVoid; (* Struct: pointer to _ecatm_foe_trfhdl *)
                                                    );

        if sFoEData.sd_retval = ECATM_OK then

          sFoEData.eSSW := _Wait4StartWriteFile; //Go on, wait for answer in next step

          sFoEData.FileSizeTransferred := 0;
          _memset(dest:=#sFoEData.FoEStatus, usByte:=0, cntr:=sizeof(sFoEData.FoEStatus));  // Reset Status as it is used in callback and my not be filled in error

          if (sFoEData.Buffer.FileSize >= sFoEData.BlockSize) then
            sFoEData.WrBlockSize := sFoEData.BlockSize;
          else
            sFoEData.WrBlockSize := sFoEData.Buffer.FileSize;
          end_if;

        elsif sFoEData.sd_retval <> ECATM_EVTC_BUSY$DINT then

          sFoEData.eSSW := t_e_FoESSW::_Error;
          HWC_LogPrintf(pThis:=this, format:="@092F (ECAT_Slave_Base::CyclicFoEHandling) Call OS_ECATM_FOE_DLD_START returned %V4", p0:=#sFoEData.sd_retval);

        end_if;

//*******************************************************************************************************************************************************
    t_e_FoESSW::_Wait4StartWriteFile:

        // Extra step os needed, wait till OS_ECATM_FOE_DLD_POLL returns ECATM_FOE_WAIT_BUFFER, then the 1st buffer must be set.
        sFoEData.sd_retval := OS_ECATM_FOE_DLD_POLL(pECAT
                                                  , ecatmhdl                                                      // ecatm   : pVoid; (* Struct: _ecatm_hdl *)
                                                  , sFoEData.pFoEHandle                                           // trfhdlp : pVoid; (* Struct: _ecatm_foe_trfhdl *)
                                                  , (sFoEData.Buffer.pFile + sFoEData.FileSizeTransferred)$^USINT  // data    : ^USINT;
                                                  , sFoEData.WrBlockSize                                          // size    : UDINT;
                                                  , #sFoEData.FoEStatus                                           // status  : pVoid; (* Struct: pointer to _ecatm_foe_status *)
                                                  );

        if sFoEData.sd_retval = ECATM_OK then

          case sFoEData.FoEStatus.state of

            ECATM_FOE_IDLE:           // transfer completed; handle freed

              sFoEData.eSSW := t_e_FoESSW::_Error;  // Error because no Files have been transferred  yet

            ECATM_FOE_DATA_READY:     // data chunk filled

              sFoEData.eSSW := _WriteFile;

            ECATM_FOE_WAIT_BUFFER:    // Ready for buffer move to next step

              sFoEData.eSSW := _WriteFile;

            ECATM_FOE_BUSY:           // FoE transfer is busy

              // Nothing to do

            ECATM_FOE_ERROR:          // FoE transfer failed; handle freed

              sFoEData.eSSW := t_e_FoESSW::_Error;
              if sFoEData.FoEStatus.error_str[0] = 0 then
                HWC_LogPrintf(pThis:=this, format:="@0930 (ECAT_Slave_Base::CyclicFoEHandling) Call OS_ECATM_FOE_DLD_POLL returned ErrorCode %V2", p0:=#sFoEData.FoEStatus.error_code);
              else
                sFoEData.FoEStatus.error_str[ECATM_FOE_MAXSTRLEN-1] := 0;   //Ensure 0 Terminaton
                HWC_LogPrintf(pThis:=this, format:="@0930 (ECAT_Slave_Base::CyclicFoEHandling) Call OS_ECATM_FOE_DLD_POLL returned ErrorCode; %V2, Error Msg: %s", p0:=#sFoEData.FoEStatus.error_code, p1:=#sFoEData.FoEStatus.error_str[0]);
              end_if;

          end_case;

        else
          sFoEData.eSSW := t_e_FoESSW::_Error;
          HWC_LogPrintf(pThis:=this, format:="@0930 (ECAT_Slave_Base::CyclicFoEHandling) Call OS_ECATM_FOE_DLD_POLL returned %d", p0:=#sFoEData.sd_retval);
        end_if;

//*******************************************************************************************************************************************************
    t_e_FoESSW::_WriteFile:

        sFoEData.sd_retval := OS_ECATM_FOE_DLD_POLL(pECAT
                                                  , ecatmhdl                                                      // ecatm   : pVoid; (* Struct: _ecatm_hdl *)
                                                  , sFoEData.pFoEHandle                                           // trfhdlp : pVoid; (* Struct: _ecatm_foe_trfhdl *)
                                                  , (sFoEData.Buffer.pFile + sFoEData.FileSizeTransferred)$^USINT  // data    : ^USINT;
                                                  , sFoEData.WrBlockSize                                          // size    : UDINT;
                                                  , #sFoEData.FoEStatus                                           // status  : pVoid; (* Struct: pointer to _ecatm_foe_status *)
                                                  );

        if sFoEData.sd_retval = ECATM_OK then

          case sFoEData.FoEStatus.state of

            ECATM_FOE_IDLE:           // transfer completed; handle freed

              sFoEData.FileSizeTransferred += sFoEData.WrBlockSize;  // Update for user Callback info
              sFoEData.eSSW := t_e_FoESSW::_Finish; //Go on

            ECATM_FOE_DATA_READY:     // data chunk filled

              // Nothing to do

            ECATM_FOE_WAIT_BUFFER:    // buffer transferred move to next

              sFoEData.FileSizeTransferred += sFoEData.WrBlockSize;
              if ((sFoEData.Buffer.FileSize - sFoEData.FileSizeTransferred) >= sFoEData.BlockSize) then
                sFoEData.WrBlockSize := sFoEData.BlockSize;
              else
                sFoEData.WrBlockSize := (sFoEData.Buffer.FileSize - sFoEData.FileSizeTransferred);
              end_if;

              // Send Update to user with new sFoEData.FileSizeTransferred
              SendFOECallback(FOEState:=BUSY);

            ECATM_FOE_BUSY:           // FoE transfer is busy

              // Nothing to do

            ECATM_FOE_ERROR:          // FoE transfer failed; handle freed

              sFoEData.eSSW := t_e_FoESSW::_Error;
              if sFoEData.FoEStatus.error_str[0] = 0 then
                HWC_LogPrintf(pThis:=this, format:="@0930 (ECAT_Slave_Base::CyclicFoEHandling) Call OS_ECATM_FOE_DLD_POLL returned ErrorCode %V2", p0:=#sFoEData.FoEStatus.error_code);
              else
                sFoEData.FoEStatus.error_str[ECATM_FOE_MAXSTRLEN-1] := 0;   //Ensure 0 Terminaton
                HWC_LogPrintf(pThis:=this, format:="@0930 (ECAT_Slave_Base::CyclicFoEHandling) Call OS_ECATM_FOE_DLD_POLL returned ErrorCode; %V2, Error Msg: %s", p0:=#sFoEData.FoEStatus.error_code, p1:=#sFoEData.FoEStatus.error_str[0]);
              end_if;

          end_case;

        else
          sFoEData.eSSW := t_e_FoESSW::_Error;
          HWC_LogPrintf(pThis:=this, format:="@0930 (ECAT_Slave_Base::CyclicFoEHandling) Call OS_ECATM_FOE_DLD_POLL returned %d", p0:=#sFoEData.sd_retval);
        end_if;

//*******************************************************************************************************************************************************
    t_e_FoESSW::_AbortFileAccess:

        sFoEData.eSSW := t_e_FoESSW::_Error;  // Should be impossible
        if sFoEData.pFoEHandle then

          sFoEData.sd_retval := OS_ECATM_FOE_ABORT( pECAT
                                                  , ecatmhdl            // ecatm   : pVoid; (* Struct: _ecatm_hdl *)
                                                  , sFoEData.pFoEHandle // trfhdlp : pVoid; (* Struct: _ecatm_foe_trfhdl *)
                                                  );
          sFoEData.eSSW := t_e_FoESSW::_Finish;
        end_if;

//*******************************************************************************************************************************************************
    t_e_FoESSW::_AbortFileAccessError:

        sFoEData.eSSW := t_e_FoESSW::_Error;  // Should be impossible
        if sFoEData.pFoEHandle then

          sFoEData.sd_retval := OS_ECATM_FOE_ABORT( pECAT
                                                  , ecatmhdl            // ecatm   : pVoid; (* Struct: _ecatm_hdl *)
                                                  , sFoEData.pFoEHandle // trfhdlp : pVoid; (* Struct: _ecatm_foe_trfhdl *)
                                                  );
          sFoEData.eSSW := t_e_FoESSW::_Error;
        end_if;

//*******************************************************************************************************************************************************
    t_e_FoESSW::_Finish:

        SendFOECallback(FOEState:=READY);

        // Reset before udIsSDOActive
        sFoEData.bFoEDataValid        := FALSE;
        sFoEData.pFoEHandle           := NIL;
        sFoEData.Buffer.pFoECallback  := NIL;
        sigclib_atomic_setU32(pValue:=#sFoEData.udIsFoEActive, value:=ECAT_SB_SDO_FREE);

        sFoEData.eSSW := t_e_FoESSW::_Idle; //Reset SSW

//*******************************************************************************************************************************************************
    t_e_FoESSW::_Error:

        SendFOECallback(FOEState:=ERROR);

        // Reset before udIsSDOActive
        sFoEData.bFoEDataValid        := FALSE;
        sFoEData.pFoEHandle           := NIL;
        sFoEData.Buffer.pFoECallback  := NIL;
        sigclib_atomic_setU32(pValue:=#sFoEData.udIsFoEActive, value:=ECAT_SB_SDO_FREE);

        sFoEData.eSSW := t_e_FoESSW::_Idle; //Reset SSW

  end_case;

END_FUNCTION

FUNCTION ECAT_Slave_Base::SendFOECallback
	VAR_INPUT
		FOEState 	: iprStates;
	END_VAR
  VAR
    UserPara  : CmdStruct;
    UserResult: Results;
  END_VAR

  if sFoEData.Buffer.pFoECallback then
    UserPara.uiCmd              := ECAT_M_FOE_CALLBACK;
    UserPara.aPara[0]           := 1;                                 //Version
    UserPara.aPara[1]$iprStates := FOEState;                          //
    UserPara.aPara[2]           := sFoEData.Buffer.ReadWriteAbortFoE; // Read or Write or arbort (0 ... Read , 1 ... Write, -1 abort)
    UserPara.aPara[3]$^CHAR     := sFoEData.Buffer.FileName;          // Filename
    UserPara.aPara[4]$UDINT     := sFoEData.FileSizeTransferred;      // FileSizeTransferred
    UserPara.aPara[5]$UDINT     := TO_UDINT(sFoEData.FoEStatus.error_code);     // Errorcode from the Slave
    sFoEData.FoEStatus.error_str[ECATM_FOE_MAXSTRLEN-1] := 0;         // Ensure 0 Terminaton
    UserPara.aPara[6]$^CHAR     := #sFoEData.FoEStatus.error_str[0];  // ErrorString from the Slave (optional)
    UserPara.aPara[7]           := sFoEData.sd_retval;                // Return code from OS Interface

    sFoEData.Buffer.pFoECallback$^VirtualBase^.NewInst(#UserPara, #UserResult);
  end_if;

END_FUNCTION

FUNCTION VIRTUAL GLOBAL ECAT_Slave_Base::StartWriteSoESSC
	VAR_INPUT
		driveno 	: DINT;
		elementflags 	: BSINT;
		IDN 	: DINT;
		pWriteData 	: ^USINT;
		udWriteLength 	: UDINT;
		udTimeout 	: UDINT;
		pCallback 	: pVoid;
	END_VAR
	VAR_OUTPUT
		retcode 	: iprStates;
	END_VAR
  VAR
    PipeSSCData : t_s_SoESSCBufferEntry;
  END_VAR

  if (pECAT^.version < ECATM_CIL_SOE_SUPPORT) then
    retcode := ERROR;
    return;
  end_if;

  //Mailbox communication is available when State is Pre-Op or higher
  if EtherCATState < ECAT_STATE_PREOP then
    retcode := ERROR;
    return;
  end_if;

  //Check input parameters
  if pWriteData = NIL then
    retcode := ERROR;
    return;
  end_if;

  if pCallback = NIL then
    retcode := ERROR;
    return;
  end_if;

  retcode := BUSY;
  // Check if pipe buffer used
  if sSSCData.pPipe then

    PipeSSCData.bWriteSSC := TRUE; //write SSC

    // Copy data to local memory before passing it to buffer
    PipeSSCData.driveno         := driveno;
    PipeSSCData.elementflags    := elementflags;
    PipeSSCData.IDN             := IDN;
    PipeSSCData.pData           := pWriteData;
    PipeSSCData.udLength        := udWriteLength;
    PipeSSCData.udTimeout       := udTimeout;
    PipeSSCData.pSSCCallback    := pCallback;

    // Add the SSC Data to buffer
    if (cPipe_Add(sSSCData.pPipe, #PipeSSCData, sizeof(t_s_SoESSCBufferEntry) ) = 1) then
      retcode := READY;
    end_if;

  // Check if currently a SSC is active, if not get lock on variables
  elsif (sigclib_atomic_cmpxchgU32(pValue:= #sSSCData.udIsSSCActive, cmpVal:=ECAT_SB_SDO_FREE, newVal:=ECAT_SB_SDO_LOCK) = ECAT_SB_SDO_FREE) then

    // Copy data to variables
    sSSCData.Buffer.bWriteSSC := TRUE; //write SSC

    sSSCData.Buffer.driveno         := driveno;
    sSSCData.Buffer.elementflags    := elementflags;
    sSSCData.Buffer.IDN             := IDN;
    sSSCData.Buffer.pData           := pWriteData;
    sSSCData.Buffer.udLength        := udWriteLength;
    sSSCData.Buffer.udTimeout       := udTimeout;
    sSSCData.Buffer.pSSCCallback    := pCallback;

    sSSCData.eSSW             := t_e_SoESSC::_StartSSCReq;

    // Set when all other data is set
    sSSCData.bSSCDataValid    := TRUE;

    retcode := READY;

  end_if;

END_FUNCTION

FUNCTION VIRTUAL GLOBAL ECAT_Slave_Base::StartReadSoESSC
	VAR_INPUT
		driveno 	: DINT;
		elementflags 	: BSINT;
		IDN 	: DINT;
		pReadData 	: ^USINT;
		udMaxDataLength 	: UDINT;
		udTimeout 	: UDINT;
		pCallback 	: pVoid;
	END_VAR
	VAR_OUTPUT
		retcode 	: iprStates;
	END_VAR
  VAR
    PipeSSCData : t_s_SoESSCBufferEntry;
  END_VAR

  if (pECAT^.version < ECATM_CIL_SOE_SUPPORT) then
    retcode := ERROR;
    return;
  end_if;

  //Mailbox communication is available when State is Pre-Op or higher
  if EtherCATState < ECAT_STATE_PREOP then
    retcode := ERROR;
    return;
  end_if;

  //Check input parameters
  if pReadData = NIL then
    retcode := ERROR;
    return;
  end_if;

  if pCallback = NIL then
    retcode := ERROR;
    return;
  end_if;

  retcode := BUSY;
  // Check if pipe buffer used
  if sSSCData.pPipe then

    // Copy data to local memory before passing it to buffer
    PipeSSCData.bWriteSSC := FALSE; //read SSC

    PipeSSCData.driveno         := driveno;
    PipeSSCData.elementflags    := elementflags;
    PipeSSCData.IDN             := IDN;
    PipeSSCData.pData           := pReadData;
    PipeSSCData.udLength        := udMaxDataLength;
    PipeSSCData.udTimeout       := udTimeout;
    PipeSSCData.pSSCCallback    := pCallback;

    // Add the SSC Data to buffer
    if (cPipe_Add(sSSCData.pPipe, #PipeSSCData, sizeof(t_s_SoESSCBufferEntry) ) = 1) then
      retcode := READY;
    end_if;

  // Check if currently a SSC is active, if not get lock on variables
  elsif (sigclib_atomic_cmpxchgU32(pValue:= #sSSCData.udIsSSCActive, cmpVal:=ECAT_SB_SDO_FREE, newVal:=ECAT_SB_SDO_LOCK) = ECAT_SB_SDO_FREE) then

    // Copy data to variables
    sSSCData.Buffer.bWriteSSC  := FALSE; //read SSC

    sSSCData.Buffer.driveno         := driveno;
    sSSCData.Buffer.elementflags    := elementflags;
    sSSCData.Buffer.IDN             := IDN;
    sSSCData.Buffer.pData           := pReadData;
    sSSCData.Buffer.udLength        := udMaxDataLength;
    sSSCData.Buffer.udTimeout       := udTimeout;
    sSSCData.Buffer.pSSCCallback    := pCallback;

    sSSCData.eSSW             := t_e_SoESSC::_StartSSCReq;

    // Set when all other data is set
    sSSCData.bSSCDataValid    := TRUE;

    retcode := READY;

  end_if;

END_FUNCTION

FUNCTION ECAT_Slave_Base::CyclicSoESSCHandling
  VAR
    UserPara  : CmdStruct;
    UserResult: Results;
  END_VAR

  if (pECAT^.version < ECATM_CIL_SOE_SUPPORT) then
    return;
  end_if;

  case sSSCData.eSSW of

//*******************************************************************************************************************************************************
    t_e_SoESSC::_StartSSCReq:  //Start SSC Request

        if (sSSCData.pPipe) &
           (sSSCData.bSSCDataValid = FALSE) then

          if cPipe_Get(pd:=#sSSCData.Buffer, p:=sSSCData.pPipe) = 1 then

            sSSCData.bSSCDataValid := TRUE;

          end_if;

        end_if;

        if sSSCData.bSSCDataValid then

          if sSSCData.Buffer.bWriteSSC = FALSE then  // Read
            //Start SSC Upload via OS
            sSSCData.sd_retval := OS_ECATM_SSC_READ_START(  pECAT
                                                          , ecatmhdl                      // ecatm           : pVoid; (* Struct: _ecatm_hdl *)
                                                          , SlaveIndex                    // slvidx          : UDINT;
                                                          , sSSCData.Buffer.driveno       // driveno         : DINT;
                                                          , sSSCData.Buffer.elementflags  // elementflags    : DINT;
                                                          , sSSCData.Buffer.IDN           // IDN             : DINT;
                                                          , sSSCData.Buffer.pData         // data            : ^USINT;    (* const *)
                                                          , sSSCData.Buffer.udLength$DINT // datamax         : DINT;
                                                          , sSSCData.Buffer.udTimeout     // tmo_ms          : UDINT;
                                                          , #sSSCData.pSSCHandle          // sschdlp         : pVoid; (* Struct: pointer to _ecatm_sschdl *)
                                                          );

          else  // Write
            //Start SSC Download via OS
            sSSCData.sd_retval := OS_ECATM_SSC_WRITE_START( pECAT
                                                          , ecatmhdl                      // ecatm           : pVoid; (* Struct: _ecatm_hdl *)
                                                          , SlaveIndex                    // slvidx          : UDINT;
                                                          , sSSCData.Buffer.driveno       // driveno         : DINT;
                                                          , sSSCData.Buffer.elementflags  // elementflags    : DINT;
                                                          , sSSCData.Buffer.IDN           // IDN             : DINT;
                                                          , sSSCData.Buffer.pData         // data            : ^USINT;    (* const *)
                                                          , sSSCData.Buffer.udLength      // datasize        : UDINT;
                                                          , sSSCData.Buffer.udTimeout     // tmo_ms          : UDINT;
                                                          , #sSSCData.pSSCHandle          // sschdlp         : pVoid; (* Struct: pointer to _ecatm_sschdl *)
                                                          );

          end_if;

          if sSSCData.sd_retval = ECATM_OK then

            sSSCData.eSSW := t_e_SoESSC::_Wait4SSCRsp; //Go on, wait for answer in next step

          elsif sSSCData.sd_retval <> ECATM_EVTC_BUSY$DINT then

            if sSSCData.Buffer.bWriteSSC = FALSE then
              HWC_LogPrintf(pThis:=this, format:="@0931 (ECAT_Slave_Base::CyclicSoESSCHandling) Call OS_ECATM_SSC_READ_START returned %d, DriveNo: %d, IDN: %d.", p0:=#sSSCData.sd_retval, p1:=#sSSCData.Buffer.driveno, p2:=#sSSCData.Buffer.IDN);
            else
              HWC_LogPrintf(pThis:=this, format:="@0932 (ECAT_Slave_Base::CyclicSoESSCHandling) Call OS_ECATM_SSC_WRITE_START returned %d, DriveNo: %d, IDN: %d.", p0:=#sSSCData.sd_retval, p1:=#sSSCData.Buffer.driveno, p2:=#sSSCData.Buffer.IDN);
            end_if;

            // Reset before udIsSDOActive
            sSSCData.bSSCDataValid    := FALSE;
            sigclib_atomic_setU32(pValue:=#sSSCData.udIsSSCActive, value:=ECAT_SB_SDO_FREE);

            if sSSCData.Buffer.pSSCCallback then
              UserPara.uiCmd          := ECAT_M_SSC_CALLBACK;
              UserPara.aPara[0]$DINT  := 1;                               // Version
              UserPara.aPara[1]$DINT  := sSSCData.sd_retval;              // Return code
              UserPara.aPara[2]$BOOL  := sSSCData.Buffer.bWriteSSC;       // Read or Write (0 ... Read , 1 ... Write)
              UserPara.aPara[3]$DINT  := sSSCData.Buffer.driveno;         // driveno
              UserPara.aPara[4]$USINT := sSSCData.Buffer.elementflags;    // elementflags
              UserPara.aPara[5]$DINT  := sSSCData.Buffer.IDN;             // IDN
              UserPara.aPara[6]$UDINT := sSSCData.Buffer.udLength;        // Datalength
              UserPara.aPara[7]$UINT  := 0;                               // SoE transfer errocode or 0 on success.

              sSSCData.Buffer.pSSCCallback$^VirtualBase^.NewInst(#UserPara, #UserResult);
            end_if;
          end_if;
        end_if;

//*******************************************************************************************************************************************************
    t_e_SoESSC::_Wait4SSCRsp:  //Receive SDO Response

      if sSSCData.Buffer.bWriteSSC = FALSE then  // Read
        sSSCData.sd_retval := OS_ECATM_SSC_READ_POLL( pECAT
                                                    , ecatmhdl                  // ecatm       : pVoid; (* Struct: _ecatm_hdl *)
                                                    , sSSCData.pSSCHandle       // sschdlp     : pVoid; (* Struct: _ecatm_sschdl *)
                                                    , #sSSCData.Buffer.udLength // datasize    : ^UDINT;
                                                    , #sSSCData.uiErrorCode     // errorcode   : ^UINT;
                                                    );
      else  // Write
        sSSCData.sd_retval := OS_ECATM_SSC_WRITE_POLL(pECAT
                                                    , ecatmhdl              // ecatm       : pVoid; (* Struct: _ecatm_hdl *)
                                                    , sSSCData.pSSCHandle   // sschdlp     : pVoid; (* Struct: _ecatm_sschdl *)
                                                    , #sSSCData.uiErrorCode // errorcode   : ^UINT;
                                                     );

      end_if;

      if sSSCData.sd_retval = ECATM_OK then

        if sSSCData.uiErrorCode <> 0 then
          sSSCData.sd_retval := -1; // Set to Not Ok if an Error code was returned
        end_if;

      elsif sSSCData.sd_retval = ECATM_EVTC_BUSY$DINT then
        return;
      else

        if sSSCData.Buffer.bWriteSSC = FALSE then
          HWC_LogPrintf(pThis:=this, format:="@0933 (ECAT_Slave_Base::CyclicSoESSCHandling) Call OS_ECATM_SSC_READ_POLL returned %d, DriveNo: %d, IDN: %d, ErrorCode: %V2.", p0:=#sSSCData.sd_retval, p1:=#sSSCData.Buffer.driveno, p2:=#sSSCData.Buffer.IDN, p3:=#sSSCData.uiErrorCode);
        else
          HWC_LogPrintf(pThis:=this, format:="@0934 (ECAT_Slave_Base::CyclicSoESSCHandling) Call OS_ECATM_SSC_WRITE_POLL returned %d, DriveNo: %d, IDN: %d, ErrorCode: %V2.", p0:=#sSSCData.sd_retval, p1:=#sSSCData.Buffer.driveno, p2:=#sSSCData.Buffer.IDN, p3:=#sSSCData.uiErrorCode);
        end_if;

      end_if;

      // Reset before udIsSDOActive
      sSSCData.bSSCDataValid    := FALSE;
      sSSCData.pSSCHandle       := NIL;   // The SDO transfer handle is invalid after a result unequal to ECATM_EVTC_BUSY was returned. (icECAT-ECATM_Reference_Manual.pdf)
      sSSCData.eSSW := t_e_SoESSC::_StartSSCReq; //Reset SSW

      sigclib_atomic_setU32(pValue:=#sSSCData.udIsSSCActive, value:=ECAT_SB_SDO_FREE);

      if sSSCData.Buffer.pSSCCallback then
        UserPara.uiCmd          := ECAT_M_SSC_CALLBACK;
        UserPara.aPara[0]$DINT  := 1;                               // Version
        UserPara.aPara[1]$DINT  := sSSCData.sd_retval;              // Return code
        UserPara.aPara[2]$BOOL  := sSSCData.Buffer.bWriteSSC;       // Read or Write (0 ... Read , 1 ... Write)
        UserPara.aPara[3]$DINT  := sSSCData.Buffer.driveno;         // driveno
        UserPara.aPara[4]$USINT := sSSCData.Buffer.elementflags;    // elementflags
        UserPara.aPara[5]$DINT  := sSSCData.Buffer.IDN;             // IDN
        UserPara.aPara[6]$UDINT := sSSCData.Buffer.udLength;        // Datalength
        UserPara.aPara[7]$UINT  := sSSCData.uiErrorCode;            // SoE transfer errocode or 0 on success.

        sSSCData.Buffer.pSSCCallback$^VirtualBase^.NewInst(#UserPara, #UserResult);
      end_if;

//*******************************************************************************************************************************************************
  end_case;

END_FUNCTION

#pragma warning(disable:73);
FUNCTION VIRTUAL ECAT_Slave_Base::AddPDOEntryFailed
	VAR_INPUT
		iErrorCode 	: DINT;
	END_VAR

  //Log Error is done in AddPDOEntry
  ClassState := _ParameterInvalid;
  EtherCATState := ECAT_STATE_NONE;

END_FUNCTION
#pragma warning(default:73);
